Fanuc KAREL source: kc00048.KL

-- PROVISIONAL review KL for V940-1; original PC SHA256 60d387081a6ce0dbc6f28720b4ae08b179a4fc1a6eaef84d6aafc5f0617fa569
-- Incomplete behavior may be omitted. Consult companion uncertainty JSON. Do not deploy.
PROGRAM KC00048
%NOLOCKGROUP
BEGIN
  -- V9_ZERO_TABLE_METADATA_HINT layout=0002_ascii; no indexed target words; source/name/runtime held
  -- UNRESOLVED_PC offsets 5-35; opcodes 27,22,22,1C,22,27,9D,31
  -- UNRESOLVED_PC offsets 40-44; opcodes 7F
END KC00048
